// TIA Portal V20 export
DATA_BLOCK "T12_Datos"   // DB48900
{ S7_Optimized_Access := 'TRUE' }
AUTHOR : IA
FAMILY : PRUEBA
VERSION : 0.1
// Tanda 7: datos
// stored: AutoNumber false
   VAR
      Arranques : DInt;   // Lo incrementa el OB100
      ErroresProg : DInt;   // Lo incrementa el OB121
      Const_Out : UInt;
      Var_Out : Int;
      Int_5 : Int := 5;
      A5 : Array[0..4] of Int;   // 1..5
      A3 : Array[1..3] of Int;   // 10,20,30
      Suma5 : DInt;
      Suma3 : DInt;
      Num5 : DInt;
      Num3 : DInt;
      Indice : Int := 7;   // Índice fuera de rango a propósito
      Error_Hecho : Bool;
   END_VAR
BEGIN
END_DATA_BLOCK
